(* IEC 61131-3 sources: codesys-framework/txt/application/WeVe Core (library)/10 Mode/Service/FB_ModeService, 12 files *)

(* ---- ActiveMode.prop.st ---- *)
PROPERTY ActiveMode : USINT

// --- BEGIN IMPLEMENTATION ---

// ----------- GET -----------
VAR
END_VAR

// -- BEGIN IMPLEMENTATION GET --
ActiveMode := _nActiveMode;

(* ---- ActiveState.prop.st ---- *)
PROPERTY ActiveState : E_ModeStates

// --- BEGIN IMPLEMENTATION ---

// ----------- GET -----------
VAR
END_VAR

// -- BEGIN IMPLEMENTATION GET --
ActiveState := _afbModes[_nActiveMode].State;

(* ---- FB_Init.method.st ---- *)
//FB_Init is always available implicitly and it is used primarily for initialization.
//The return value is not evaluated. For a specific influence, you can also declare the
//methods explicitly and provide additional code there with the standard initialization
//code. You can evaluate the return value.
METHOD FB_Init: BOOL
VAR_INPUT
    bInitRetains: BOOL; // TRUE: the retain variables are initialized (reset warm / reset cold)
    bInCopyCode: BOOL;  // TRUE: the instance will be copied to the copy code afterward (online change)

	fbEventSrv 				: I_EventService;
	fbLogger 				: I_Logger;
	fbEvents 				: I_EventGroup;		// de gedeelde FB_ModeEventGroup, mag 0 zijn
	afbModes 				: ARRAY[0..cNbrOfModes] OF I_Mode;
END_VAR

// --- BEGIN IMPLEMENTATION ---

_fbEventSrv := fbEventSrv;
_fbLogger := fbLogger;
_fbEvents := fbEvents;
_afbModes := afbModes;

_xInit := TRUE;

(* ---- Init.method.st ---- *)
METHOD PRIVATE Init
VAR_INPUT
END_VAR
VAR
	i 	: USINT;
END_VAR

// --- BEGIN IMPLEMENTATION ---

FOR i := 0 TO cNbrOfModes DO

	IF _afbModes[i] <> 0 THEN
		_afbModes[i].Active := i = _nActiveMode;
	END_IF

END_FOR

(* ---- Initialize.method.st ---- *)
METHOD Initialize
VAR_INPUT
END_VAR

// --- BEGIN IMPLEMENTATION ---

_nActiveMode := E_DefaultModes.Auto;

IF _afbModes[_nActiveMode] <> 0 THEN
	_afbModes[_nActiveMode].State := E_ModeStates.Off;
END_IF

(* ---- RequestMode.method.st ---- *)
METHOD RequestMode
VAR_INPUT
	nMode		: USINT;
END_VAR
VAR
	i 			: USINT;
	scPayload 	: SC_EventPayload;
END_VAR

// --- BEGIN IMPLEMENTATION ---

IF _afbModes[nMode] = 0 THEN
	RETURN;
END_IF

scPayload.asPayload[0] := _afbModes[nMode].Name;

IF _fbEvents <> 0 THEN
	_fbEvents.Log(iEvent := E_ModeEvents.ModeRequest, scPayload := scPayload);
END_IF

IF _afbModes[_nActiveMode].State = E_ModeStates.Standby THEN

	FOR i := 0 TO cNbrOfModes DO

		IF _afbModes[i] <> 0 THEN
			_afbModes[i].State := E_ModeStates.Off;
		END_IF

	END_FOR

	_nActiveMode := nMode;
	_afbModes[nMode].Active := TRUE;

ELSIF _fbEvents <> 0 THEN

	_fbEvents.Log(iEvent := E_ModeEvents.ModeRequestInvalid, scPayload := scPayload);

END_IF

(* ---- ResetEvents.method.st ---- *)
METHOD ResetEvents : BOOL

// --- BEGIN IMPLEMENTATION ---

IF _afbModes[_nActiveMode] <> 0 THEN
	_afbModes[_nActiveMode].ResetEvents();
END_IF

(* ---- ResetMachine.method.st ---- *)
METHOD ResetMachine : BOOL

// --- BEGIN IMPLEMENTATION ---

IF _afbModes[_nActiveMode] <> 0 THEN
	_afbModes[_nActiveMode].ResetMachine();
END_IF

(* ---- ResetSafety.method.st ---- *)
METHOD ResetSafety : BOOL

// --- BEGIN IMPLEMENTATION ---

IF _afbModes[_nActiveMode] <> 0 THEN
	_afbModes[_nActiveMode].ResetSafety();
END_IF

(* ---- StartRequest.method.st ---- *)
METHOD StartRequest

// --- BEGIN IMPLEMENTATION ---

IF _afbModes[_nActiveMode] <> 0 THEN
	_afbModes[_nActiveMode].StartRequest();
END_IF

(* ---- StopRequest.method.st ---- *)
METHOD StopRequest

// --- BEGIN IMPLEMENTATION ---

IF _afbModes[_nActiveMode] <> 0 THEN
	_afbModes[_nActiveMode].StopRequest();
END_IF

(* ---- UserRequest.method.st ---- *)
METHOD UserRequest
VAR_INPUT
	nRequest	: UINT;
	pData		: POINTER TO ARRAY [0..255] OF BYTE := 0;
	pSize		: ULINT := 0;
END_VAR

// --- BEGIN IMPLEMENTATION ---

IF _afbModes[_nActiveMode] <> 0 THEN
	_afbModes[_nActiveMode].UserRequest(nRequest := nRequest, pData := pData,  pSize := pSize);
END_IF
